Staubli VAL3: setAnaOutput.pgx

public program setAnaOutput(aio& x_aOut, num x_nValue, bool& x_bError)
  local string l_sDesc
  local string l_sPath
begin
  if ioStatus(x_aOut,l_sDesc,l_sPath)>=0
    x_bError=false
    aioSet(x_aOut,x_nValue)
  else
    x_bError=true
//    logMsg("Signal "+l_sPath+" error."+"Description:"+l_sDesc)
  endIf
end
